(* IEC 61131-3 sources: STAR-PLC-Agent/results/raw/four_group_20261114/star_terra/PUB012/generation/sim_00, 1 file *)

(* ---- test_program.st ---- *)
PROGRAM PLC_PRG
VAR
 BenchStep : UDINT := 0;
 BenchCalls : UDINT := 0;
 BenchDone : BOOL := FALSE;
 BenchLastTime : TIME := T#0ms;
 BenchClockReady : BOOL := FALSE;
 BenchCurrentTime : TIME := T#0ms;
 TraceDt : ARRAY[0..15] OF UDINT;
 BenchUut0 : FB_Task;
 BenchUut1 : FB_Task;
 TraceIn_THICKNESS_FAULT : ARRAY[0..15] OF BOOL;
 TraceIn_THICKNESS_SIGNAL_VALID : ARRAY[0..15] OF BOOL;
 TraceIn_CUTTING_RUN : ARRAY[0..15] OF BOOL;
 TraceIn_FaultTimestamp : ARRAY[0..15] OF DINT;
 TraceIn_CycleTime : ARRAY[0..15] OF TIME;
 TraceOut_THICKNESS_ALARM : ARRAY[0..15] OF BOOL;
 TraceOut_Slab_Fault_Counter : ARRAY[0..15] OF UINT;
 TraceOut_Slab_Runtime_Accumulator : ARRAY[0..15] OF LTIME;
 TraceOut_Slab_Fault_History_0 : ARRAY[0..15] OF DINT;
 TraceOut_Slab_Fault_History_1 : ARRAY[0..15] OF DINT;
 TraceOut_Slab_Fault_History_2 : ARRAY[0..15] OF DINT;
 TraceOut_Slab_Fault_History_3 : ARRAY[0..15] OF DINT;
 TraceOut_Slab_Fault_History_4 : ARRAY[0..15] OF DINT;
END_VAR

IF NOT BenchDone THEN
 BenchCurrentTime := TIME();
 IF NOT BenchClockReady THEN
  BenchLastTime := BenchCurrentTime;
  BenchClockReady := TRUE;
 ELSE
 CASE BenchStep OF
 0:
  IF BenchCurrentTime - BenchLastTime >= UDINT_TO_TIME(10) THEN
   TraceDt[0] := TIME_TO_UDINT(BenchCurrentTime - BenchLastTime);
   BenchLastTime := BenchCurrentTime;
   BenchUut0.THICKNESS_FAULT := FALSE;
   BenchUut0.THICKNESS_SIGNAL_VALID := FALSE;
   BenchUut0.CUTTING_RUN := TRUE;
   BenchUut0.FaultTimestamp := DINT#0;
   BenchUut0.CycleTime := TIME#10ms;
   TraceIn_THICKNESS_FAULT[0] := BenchUut0.THICKNESS_FAULT;
   TraceIn_THICKNESS_SIGNAL_VALID[0] := BenchUut0.THICKNESS_SIGNAL_VALID;
   TraceIn_CUTTING_RUN[0] := BenchUut0.CUTTING_RUN;
   TraceIn_FaultTimestamp[0] := BenchUut0.FaultTimestamp;
   TraceIn_CycleTime[0] := BenchUut0.CycleTime;
   BenchUut0();
   TraceOut_THICKNESS_ALARM[0] := BenchUut0.THICKNESS_ALARM;
   TraceOut_Slab_Fault_Counter[0] := BenchUut0.Slab_Fault_Counter;
   TraceOut_Slab_Runtime_Accumulator[0] := BenchUut0.Slab_Runtime_Accumulator;
   TraceOut_Slab_Fault_History_0[0] := BenchUut0.Slab_Fault_History[0];
   TraceOut_Slab_Fault_History_1[0] := BenchUut0.Slab_Fault_History[1];
   TraceOut_Slab_Fault_History_2[0] := BenchUut0.Slab_Fault_History[2];
   TraceOut_Slab_Fault_History_3[0] := BenchUut0.Slab_Fault_History[3];
   TraceOut_Slab_Fault_History_4[0] := BenchUut0.Slab_Fault_History[4];
   BenchCalls := BenchCalls + 1;
   BenchStep := BenchStep + 1;
  END_IF;
 1:
  IF BenchCurrentTime - BenchLastTime >= UDINT_TO_TIME(100) THEN
   TraceDt[1] := TIME_TO_UDINT(BenchCurrentTime - BenchLastTime);
   BenchLastTime := BenchCurrentTime;
   BenchUut0.THICKNESS_FAULT := FALSE;
   BenchUut0.THICKNESS_SIGNAL_VALID := TRUE;
   BenchUut0.CUTTING_RUN := TRUE;
   BenchUut0.FaultTimestamp := DINT#0;
   BenchUut0.CycleTime := TIME#100ms;
   TraceIn_THICKNESS_FAULT[1] := BenchUut0.THICKNESS_FAULT;
   TraceIn_THICKNESS_SIGNAL_VALID[1] := BenchUut0.THICKNESS_SIGNAL_VALID;
   TraceIn_CUTTING_RUN[1] := BenchUut0.CUTTING_RUN;
   TraceIn_FaultTimestamp[1] := BenchUut0.FaultTimestamp;
   TraceIn_CycleTime[1] := BenchUut0.CycleTime;
   BenchUut0();
   TraceOut_THICKNESS_ALARM[1] := BenchUut0.THICKNESS_ALARM;
   TraceOut_Slab_Fault_Counter[1] := BenchUut0.Slab_Fault_Counter;
   TraceOut_Slab_Runtime_Accumulator[1] := BenchUut0.Slab_Runtime_Accumulator;
   TraceOut_Slab_Fault_History_0[1] := BenchUut0.Slab_Fault_History[0];
   TraceOut_Slab_Fault_History_1[1] := BenchUut0.Slab_Fault_History[1];
   TraceOut_Slab_Fault_History_2[1] := BenchUut0.Slab_Fault_History[2];
   TraceOut_Slab_Fault_History_3[1] := BenchUut0.Slab_Fault_History[3];
   TraceOut_Slab_Fault_History_4[1] := BenchUut0.Slab_Fault_History[4];
   BenchCalls := BenchCalls + 1;
   BenchStep := BenchStep + 1;
  END_IF;
 2:
  IF BenchCurrentTime - BenchLastTime >= UDINT_TO_TIME(20) THEN
   TraceDt[2] := TIME_TO_UDINT(BenchCurrentTime - BenchLastTime);
   BenchLastTime := BenchCurrentTime;
   BenchUut0.THICKNESS_FAULT := TRUE;
   BenchUut0.THICKNESS_SIGNAL_VALID := TRUE;
   BenchUut0.CUTTING_RUN := TRUE;
   BenchUut0.FaultTimestamp := DINT#101;
   BenchUut0.CycleTime := TIME#20ms;
   TraceIn_THICKNESS_FAULT[2] := BenchUut0.THICKNESS_FAULT;
   TraceIn_THICKNESS_SIGNAL_VALID[2] := BenchUut0.THICKNESS_SIGNAL_VALID;
   TraceIn_CUTTING_RUN[2] := BenchUut0.CUTTING_RUN;
   TraceIn_FaultTimestamp[2] := BenchUut0.FaultTimestamp;
   TraceIn_CycleTime[2] := BenchUut0.CycleTime;
   BenchUut0();
   TraceOut_THICKNESS_ALARM[2] := BenchUut0.THICKNESS_ALARM;
   TraceOut_Slab_Fault_Counter[2] := BenchUut0.Slab_Fault_Counter;
   TraceOut_Slab_Runtime_Accumulator[2] := BenchUut0.Slab_Runtime_Accumulator;
   TraceOut_Slab_Fault_History_0[2] := BenchUut0.Slab_Fault_History[0];
   TraceOut_Slab_Fault_History_1[2] := BenchUut0.Slab_Fault_History[1];
   TraceOut_Slab_Fault_History_2[2] := BenchUut0.Slab_Fault_History[2];
   TraceOut_Slab_Fault_History_3[2] := BenchUut0.Slab_Fault_History[3];
   TraceOut_Slab_Fault_History_4[2] := BenchUut0.Slab_Fault_History[4];
   BenchCalls := BenchCalls + 1;
   BenchStep := BenchStep + 1;
  END_IF;
 3:
  IF BenchCurrentTime - BenchLastTime >= UDINT_TO_TIME(600) THEN
   TraceDt[3] := TIME_TO_UDINT(BenchCurrentTime - BenchLastTime);
   BenchLastTime := BenchCurrentTime;
   BenchUut0.THICKNESS_FAULT := TRUE;
   BenchUut0.THICKNESS_SIGNAL_VALID := TRUE;
   BenchUut0.CUTTING_RUN := TRUE;
   BenchUut0.FaultTimestamp := DINT#999;
   BenchUut0.CycleTime := TIME#600ms;
   TraceIn_THICKNESS_FAULT[3] := BenchUut0.THICKNESS_FAULT;
   TraceIn_THICKNESS_SIGNAL_VALID[3] := BenchUut0.THICKNESS_SIGNAL_VALID;
   TraceIn_CUTTING_RUN[3] := BenchUut0.CUTTING_RUN;
   TraceIn_FaultTimestamp[3] := BenchUut0.FaultTimestamp;
   TraceIn_CycleTime[3] := BenchUut0.CycleTime;
   BenchUut0();
   TraceOut_THICKNESS_ALARM[3] := BenchUut0.THICKNESS_ALARM;
   TraceOut_Slab_Fault_Counter[3] := BenchUut0.Slab_Fault_Counter;
   TraceOut_Slab_Runtime_Accumulator[3] := BenchUut0.Slab_Runtime_Accumulator;
   TraceOut_Slab_Fault_History_0[3] := BenchUut0.Slab_Fault_History[0];
   TraceOut_Slab_Fault_History_1[3] := BenchUut0.Slab_Fault_History[1];
   TraceOut_Slab_Fault_History_2[3] := BenchUut0.Slab_Fault_History[2];
   TraceOut_Slab_Fault_History_3[3] := BenchUut0.Slab_Fault_History[3];
   TraceOut_Slab_Fault_History_4[3] := BenchUut0.Slab_Fault_History[4];
   BenchCalls := BenchCalls + 1;
   BenchStep := BenchStep + 1;
  END_IF;
 4:
  IF BenchCurrentTime - BenchLastTime >= UDINT_TO_TIME(1) THEN
   TraceDt[4] := TIME_TO_UDINT(BenchCurrentTime - BenchLastTime);
   BenchLastTime := BenchCurrentTime;
   BenchUut0.THICKNESS_FAULT := FALSE;
   BenchUut0.THICKNESS_SIGNAL_VALID := TRUE;
   BenchUut0.CUTTING_RUN := FALSE;
   BenchUut0.FaultTimestamp := DINT#999;
   BenchUut0.CycleTime := TIME#1ms;
   TraceIn_THICKNESS_FAULT[4] := BenchUut0.THICKNESS_FAULT;
   TraceIn_THICKNESS_SIGNAL_VALID[4] := BenchUut0.THICKNESS_SIGNAL_VALID;
   TraceIn_CUTTING_RUN[4] := BenchUut0.CUTTING_RUN;
   TraceIn_FaultTimestamp[4] := BenchUut0.FaultTimestamp;
   TraceIn_CycleTime[4] := BenchUut0.CycleTime;
   BenchUut0();
   TraceOut_THICKNESS_ALARM[4] := BenchUut0.THICKNESS_ALARM;
   TraceOut_Slab_Fault_Counter[4] := BenchUut0.Slab_Fault_Counter;
   TraceOut_Slab_Runtime_Accumulator[4] := BenchUut0.Slab_Runtime_Accumulator;
   TraceOut_Slab_Fault_History_0[4] := BenchUut0.Slab_Fault_History[0];
   TraceOut_Slab_Fault_History_1[4] := BenchUut0.Slab_Fault_History[1];
   TraceOut_Slab_Fault_History_2[4] := BenchUut0.Slab_Fault_History[2];
   TraceOut_Slab_Fault_History_3[4] := BenchUut0.Slab_Fault_History[3];
   TraceOut_Slab_Fault_History_4[4] := BenchUut0.Slab_Fault_History[4];
   BenchCalls := BenchCalls + 1;
   BenchStep := BenchStep + 1;
  END_IF;
 5:
  IF BenchCurrentTime - BenchLastTime >= UDINT_TO_TIME(20) THEN
   TraceDt[5] := TIME_TO_UDINT(BenchCurrentTime - BenchLastTime);
   BenchLastTime := BenchCurrentTime;
   BenchUut0.THICKNESS_FAULT := TRUE;
   BenchUut0.THICKNESS_SIGNAL_VALID := TRUE;
   BenchUut0.CUTTING_RUN := TRUE;
   BenchUut0.FaultTimestamp := DINT#202;
   BenchUut0.CycleTime := TIME#20ms;
   TraceIn_THICKNESS_FAULT[5] := BenchUut0.THICKNESS_FAULT;
   TraceIn_THICKNESS_SIGNAL_VALID[5] := BenchUut0.THICKNESS_SIGNAL_VALID;
   TraceIn_CUTTING_RUN[5] := BenchUut0.CUTTING_RUN;
   TraceIn_FaultTimestamp[5] := BenchUut0.FaultTimestamp;
   TraceIn_CycleTime[5] := BenchUut0.CycleTime;
   BenchUut0();
   TraceOut_THICKNESS_ALARM[5] := BenchUut0.THICKNESS_ALARM;
   TraceOut_Slab_Fault_Counter[5] := BenchUut0.Slab_Fault_Counter;
   TraceOut_Slab_Runtime_Accumulator[5] := BenchUut0.Slab_Runtime_Accumulator;
   TraceOut_Slab_Fault_History_0[5] := BenchUut0.Slab_Fault_History[0];
   TraceOut_Slab_Fault_History_1[5] := BenchUut0.Slab_Fault_History[1];
   TraceOut_Slab_Fault_History_2[5] := BenchUut0.Slab_Fault_History[2];
   TraceOut_Slab_Fault_History_3[5] := BenchUut0.Slab_Fault_History[3];
   TraceOut_Slab_Fault_History_4[5] := BenchUut0.Slab_Fault_History[4];
   BenchCalls := BenchCalls + 1;
   BenchStep := BenchStep + 1;
  END_IF;
 6:
  IF BenchCurrentTime - BenchLastTime >= UDINT_TO_TIME(10) THEN
   TraceDt[6] := TIME_TO_UDINT(BenchCurrentTime - BenchLastTime);
   BenchLastTime := BenchCurrentTime;
   BenchUut0.THICKNESS_FAULT := TRUE;
   BenchUut0.THICKNESS_SIGNAL_VALID := FALSE;
   BenchUut0.CUTTING_RUN := TRUE;
   BenchUut0.FaultTimestamp := DINT#250;
   BenchUut0.CycleTime := TIME#10ms;
   TraceIn_THICKNESS_FAULT[6] := BenchUut0.THICKNESS_FAULT;
   TraceIn_THICKNESS_SIGNAL_VALID[6] := BenchUut0.THICKNESS_SIGNAL_VALID;
   TraceIn_CUTTING_RUN[6] := BenchUut0.CUTTING_RUN;
   TraceIn_FaultTimestamp[6] := BenchUut0.FaultTimestamp;
   TraceIn_CycleTime[6] := BenchUut0.CycleTime;
   BenchUut0();
   TraceOut_THICKNESS_ALARM[6] := BenchUut0.THICKNESS_ALARM;
   TraceOut_Slab_Fault_Counter[6] := BenchUut0.Slab_Fault_Counter;
   TraceOut_Slab_Runtime_Accumulator[6] := BenchUut0.Slab_Runtime_Accumulator;
   TraceOut_Slab_Fault_History_0[6] := BenchUut0.Slab_Fault_History[0];
   TraceOut_Slab_Fault_History_1[6] := BenchUut0.Slab_Fault_History[1];
   TraceOut_Slab_Fault_History_2[6] := BenchUut0.Slab_Fault_History[2];
   TraceOut_Slab_Fault_History_3[6] := BenchUut0.Slab_Fault_History[3];
   TraceOut_Slab_Fault_History_4[6] := BenchUut0.Slab_Fault_History[4];
   BenchCalls := BenchCalls + 1;
   BenchStep := BenchStep + 1;
  END_IF;
 7:
  IF BenchCurrentTime - BenchLastTime >= UDINT_TO_TIME(10) THEN
   TraceDt[7] := TIME_TO_UDINT(BenchCurrentTime - BenchLastTime);
   BenchLastTime := BenchCurrentTime;
   BenchUut0.THICKNESS_FAULT := TRUE;
   BenchUut0.THICKNESS_SIGNAL_VALID := TRUE;
   BenchUut0.CUTTING_RUN := TRUE;
   BenchUut0.FaultTimestamp := DINT#303;
   BenchUut0.CycleTime := TIME#10ms;
   TraceIn_THICKNESS_FAULT[7] := BenchUut0.THICKNESS_FAULT;
   TraceIn_THICKNESS_SIGNAL_VALID[7] := BenchUut0.THICKNESS_SIGNAL_VALID;
   TraceIn_CUTTING_RUN[7] := BenchUut0.CUTTING_RUN;
   TraceIn_FaultTimestamp[7] := BenchUut0.FaultTimestamp;
   TraceIn_CycleTime[7] := BenchUut0.CycleTime;
   BenchUut0();
   TraceOut_THICKNESS_ALARM[7] := BenchUut0.THICKNESS_ALARM;
   TraceOut_Slab_Fault_Counter[7] := BenchUut0.Slab_Fault_Counter;
   TraceOut_Slab_Runtime_Accumulator[7] := BenchUut0.Slab_Runtime_Accumulator;
   TraceOut_Slab_Fault_History_0[7] := BenchUut0.Slab_Fault_History[0];
   TraceOut_Slab_Fault_History_1[7] := BenchUut0.Slab_Fault_History[1];
   TraceOut_Slab_Fault_History_2[7] := BenchUut0.Slab_Fault_History[2];
   TraceOut_Slab_Fault_History_3[7] := BenchUut0.Slab_Fault_History[3];
   TraceOut_Slab_Fault_History_4[7] := BenchUut0.Slab_Fault_History[4];
   BenchCalls := BenchCalls + 1;
   BenchStep := BenchStep + 1;
  END_IF;
 8:
  IF BenchCurrentTime - BenchLastTime >= UDINT_TO_TIME(1) THEN
   TraceDt[8] := TIME_TO_UDINT(BenchCurrentTime - BenchLastTime);
   BenchLastTime := BenchCurrentTime;
   BenchUut1.THICKNESS_FAULT := FALSE;
   BenchUut1.THICKNESS_SIGNAL_VALID := TRUE;
   BenchUut1.CUTTING_RUN := TRUE;
   BenchUut1.FaultTimestamp := DINT#0;
   BenchUut1.CycleTime := TIME#1ms;
   TraceIn_THICKNESS_FAULT[8] := BenchUut1.THICKNESS_FAULT;
   TraceIn_THICKNESS_SIGNAL_VALID[8] := BenchUut1.THICKNESS_SIGNAL_VALID;
   TraceIn_CUTTING_RUN[8] := BenchUut1.CUTTING_RUN;
   TraceIn_FaultTimestamp[8] := BenchUut1.FaultTimestamp;
   TraceIn_CycleTime[8] := BenchUut1.CycleTime;
   BenchUut1();
   TraceOut_THICKNESS_ALARM[8] := BenchUut1.THICKNESS_ALARM;
   TraceOut_Slab_Fault_Counter[8] := BenchUut1.Slab_Fault_Counter;
   TraceOut_Slab_Runtime_Accumulator[8] := BenchUut1.Slab_Runtime_Accumulator;
   TraceOut_Slab_Fault_History_0[8] := BenchUut1.Slab_Fault_History[0];
   TraceOut_Slab_Fault_History_1[8] := BenchUut1.Slab_Fault_History[1];
   TraceOut_Slab_Fault_History_2[8] := BenchUut1.Slab_Fault_History[2];
   TraceOut_Slab_Fault_History_3[8] := BenchUut1.Slab_Fault_History[3];
   TraceOut_Slab_Fault_History_4[8] := BenchUut1.Slab_Fault_History[4];
   BenchCalls := BenchCalls + 1;
   BenchStep := BenchStep + 1;
  END_IF;
 9:
  IF BenchCurrentTime - BenchLastTime >= UDINT_TO_TIME(1) THEN
   TraceDt[9] := TIME_TO_UDINT(BenchCurrentTime - BenchLastTime);
   BenchLastTime := BenchCurrentTime;
   BenchUut1.THICKNESS_FAULT := TRUE;
   BenchUut1.THICKNESS_SIGNAL_VALID := TRUE;
   BenchUut1.CUTTING_RUN := TRUE;
   BenchUut1.FaultTimestamp := DINT#-2147483648;
   BenchUut1.CycleTime := TIME#1ms;
   TraceIn_THICKNESS_FAULT[9] := BenchUut1.THICKNESS_FAULT;
   TraceIn_THICKNESS_SIGNAL_VALID[9] := BenchUut1.THICKNESS_SIGNAL_VALID;
   TraceIn_CUTTING_RUN[9] := BenchUut1.CUTTING_RUN;
   TraceIn_FaultTimestamp[9] := BenchUut1.FaultTimestamp;
   TraceIn_CycleTime[9] := BenchUut1.CycleTime;
   BenchUut1();
   TraceOut_THICKNESS_ALARM[9] := BenchUut1.THICKNESS_ALARM;
   TraceOut_Slab_Fault_Counter[9] := BenchUut1.Slab_Fault_Counter;
   TraceOut_Slab_Runtime_Accumulator[9] := BenchUut1.Slab_Runtime_Accumulator;
   TraceOut_Slab_Fault_History_0[9] := BenchUut1.Slab_Fault_History[0];
   TraceOut_Slab_Fault_History_1[9] := BenchUut1.Slab_Fault_History[1];
   TraceOut_Slab_Fault_History_2[9] := BenchUut1.Slab_Fault_History[2];
   TraceOut_Slab_Fault_History_3[9] := BenchUut1.Slab_Fault_History[3];
   TraceOut_Slab_Fault_History_4[9] := BenchUut1.Slab_Fault_History[4];
   BenchCalls := BenchCalls + 1;
   BenchStep := BenchStep + 1;
  END_IF;
 10:
  IF BenchCurrentTime - BenchLastTime >= UDINT_TO_TIME(499) THEN
   TraceDt[10] := TIME_TO_UDINT(BenchCurrentTime - BenchLastTime);
   BenchLastTime := BenchCurrentTime;
   BenchUut1.THICKNESS_FAULT := FALSE;
   BenchUut1.THICKNESS_SIGNAL_VALID := TRUE;
   BenchUut1.CUTTING_RUN := TRUE;
   BenchUut1.FaultTimestamp := DINT#0;
   BenchUut1.CycleTime := TIME#499ms;
   TraceIn_THICKNESS_FAULT[10] := BenchUut1.THICKNESS_FAULT;
   TraceIn_THICKNESS_SIGNAL_VALID[10] := BenchUut1.THICKNESS_SIGNAL_VALID;
   TraceIn_CUTTING_RUN[10] := BenchUut1.CUTTING_RUN;
   TraceIn_FaultTimestamp[10] := BenchUut1.FaultTimestamp;
   TraceIn_CycleTime[10] := BenchUut1.CycleTime;
   BenchUut1();
   TraceOut_THICKNESS_ALARM[10] := BenchUut1.THICKNESS_ALARM;
   TraceOut_Slab_Fault_Counter[10] := BenchUut1.Slab_Fault_Counter;
   TraceOut_Slab_Runtime_Accumulator[10] := BenchUut1.Slab_Runtime_Accumulator;
   TraceOut_Slab_Fault_History_0[10] := BenchUut1.Slab_Fault_History[0];
   TraceOut_Slab_Fault_History_1[10] := BenchUut1.Slab_Fault_History[1];
   TraceOut_Slab_Fault_History_2[10] := BenchUut1.Slab_Fault_History[2];
   TraceOut_Slab_Fault_History_3[10] := BenchUut1.Slab_Fault_History[3];
   TraceOut_Slab_Fault_History_4[10] := BenchUut1.Slab_Fault_History[4];
   BenchCalls := BenchCalls + 1;
   BenchStep := BenchStep + 1;
  END_IF;
 11:
  IF BenchCurrentTime - BenchLastTime >= UDINT_TO_TIME(1) THEN
   TraceDt[11] := TIME_TO_UDINT(BenchCurrentTime - BenchLastTime);
   BenchLastTime := BenchCurrentTime;
   BenchUut1.THICKNESS_FAULT := TRUE;
   BenchUut1.THICKNESS_SIGNAL_VALID := TRUE;
   BenchUut1.CUTTING_RUN := TRUE;
   BenchUut1.FaultTimestamp := DINT#2147483647;
   BenchUut1.CycleTime := TIME#1ms;
   TraceIn_THICKNESS_FAULT[11] := BenchUut1.THICKNESS_FAULT;
   TraceIn_THICKNESS_SIGNAL_VALID[11] := BenchUut1.THICKNESS_SIGNAL_VALID;
   TraceIn_CUTTING_RUN[11] := BenchUut1.CUTTING_RUN;
   TraceIn_FaultTimestamp[11] := BenchUut1.FaultTimestamp;
   TraceIn_CycleTime[11] := BenchUut1.CycleTime;
   BenchUut1();
   TraceOut_THICKNESS_ALARM[11] := BenchUut1.THICKNESS_ALARM;
   TraceOut_Slab_Fault_Counter[11] := BenchUut1.Slab_Fault_Counter;
   TraceOut_Slab_Runtime_Accumulator[11] := BenchUut1.Slab_Runtime_Accumulator;
   TraceOut_Slab_Fault_History_0[11] := BenchUut1.Slab_Fault_History[0];
   TraceOut_Slab_Fault_History_1[11] := BenchUut1.Slab_Fault_History[1];
   TraceOut_Slab_Fault_History_2[11] := BenchUut1.Slab_Fault_History[2];
   TraceOut_Slab_Fault_History_3[11] := BenchUut1.Slab_Fault_History[3];
   TraceOut_Slab_Fault_History_4[11] := BenchUut1.Slab_Fault_History[4];
   BenchCalls := BenchCalls + 1;
   BenchStep := BenchStep + 1;
  END_IF;
 12:
  IF BenchCurrentTime - BenchLastTime >= UDINT_TO_TIME(499) THEN
   TraceDt[12] := TIME_TO_UDINT(BenchCurrentTime - BenchLastTime);
   BenchLastTime := BenchCurrentTime;
   BenchUut1.THICKNESS_FAULT := FALSE;
   BenchUut1.THICKNESS_SIGNAL_VALID := TRUE;
   BenchUut1.CUTTING_RUN := TRUE;
   BenchUut1.FaultTimestamp := DINT#0;
   BenchUut1.CycleTime := TIME#499ms;
   TraceIn_THICKNESS_FAULT[12] := BenchUut1.THICKNESS_FAULT;
   TraceIn_THICKNESS_SIGNAL_VALID[12] := BenchUut1.THICKNESS_SIGNAL_VALID;
   TraceIn_CUTTING_RUN[12] := BenchUut1.CUTTING_RUN;
   TraceIn_FaultTimestamp[12] := BenchUut1.FaultTimestamp;
   TraceIn_CycleTime[12] := BenchUut1.CycleTime;
   BenchUut1();
   TraceOut_THICKNESS_ALARM[12] := BenchUut1.THICKNESS_ALARM;
   TraceOut_Slab_Fault_Counter[12] := BenchUut1.Slab_Fault_Counter;
   TraceOut_Slab_Runtime_Accumulator[12] := BenchUut1.Slab_Runtime_Accumulator;
   TraceOut_Slab_Fault_History_0[12] := BenchUut1.Slab_Fault_History[0];
   TraceOut_Slab_Fault_History_1[12] := BenchUut1.Slab_Fault_History[1];
   TraceOut_Slab_Fault_History_2[12] := BenchUut1.Slab_Fault_History[2];
   TraceOut_Slab_Fault_History_3[12] := BenchUut1.Slab_Fault_History[3];
   TraceOut_Slab_Fault_History_4[12] := BenchUut1.Slab_Fault_History[4];
   BenchCalls := BenchCalls + 1;
   BenchStep := BenchStep + 1;
  END_IF;
 13:
  IF BenchCurrentTime - BenchLastTime >= UDINT_TO_TIME(1) THEN
   TraceDt[13] := TIME_TO_UDINT(BenchCurrentTime - BenchLastTime);
   BenchLastTime := BenchCurrentTime;
   BenchUut1.THICKNESS_FAULT := FALSE;
   BenchUut1.THICKNESS_SIGNAL_VALID := TRUE;
   BenchUut1.CUTTING_RUN := TRUE;
   BenchUut1.FaultTimestamp := DINT#0;
   BenchUut1.CycleTime := TIME#1ms;
   TraceIn_THICKNESS_FAULT[13] := BenchUut1.THICKNESS_FAULT;
   TraceIn_THICKNESS_SIGNAL_VALID[13] := BenchUut1.THICKNESS_SIGNAL_VALID;
   TraceIn_CUTTING_RUN[13] := BenchUut1.CUTTING_RUN;
   TraceIn_FaultTimestamp[13] := BenchUut1.FaultTimestamp;
   TraceIn_CycleTime[13] := BenchUut1.CycleTime;
   BenchUut1();
   TraceOut_THICKNESS_ALARM[13] := BenchUut1.THICKNESS_ALARM;
   TraceOut_Slab_Fault_Counter[13] := BenchUut1.Slab_Fault_Counter;
   TraceOut_Slab_Runtime_Accumulator[13] := BenchUut1.Slab_Runtime_Accumulator;
   TraceOut_Slab_Fault_History_0[13] := BenchUut1.Slab_Fault_History[0];
   TraceOut_Slab_Fault_History_1[13] := BenchUut1.Slab_Fault_History[1];
   TraceOut_Slab_Fault_History_2[13] := BenchUut1.Slab_Fault_History[2];
   TraceOut_Slab_Fault_History_3[13] := BenchUut1.Slab_Fault_History[3];
   TraceOut_Slab_Fault_History_4[13] := BenchUut1.Slab_Fault_History[4];
   BenchCalls := BenchCalls + 1;
   BenchStep := BenchStep + 1;
  END_IF;
 14:
  IF BenchCurrentTime - BenchLastTime >= UDINT_TO_TIME(1) THEN
   TraceDt[14] := TIME_TO_UDINT(BenchCurrentTime - BenchLastTime);
   BenchLastTime := BenchCurrentTime;
   BenchUut1.THICKNESS_FAULT := TRUE;
   BenchUut1.THICKNESS_SIGNAL_VALID := TRUE;
   BenchUut1.CUTTING_RUN := TRUE;
   BenchUut1.FaultTimestamp := DINT#0;
   BenchUut1.CycleTime := TIME#1ms;
   TraceIn_THICKNESS_FAULT[14] := BenchUut1.THICKNESS_FAULT;
   TraceIn_THICKNESS_SIGNAL_VALID[14] := BenchUut1.THICKNESS_SIGNAL_VALID;
   TraceIn_CUTTING_RUN[14] := BenchUut1.CUTTING_RUN;
   TraceIn_FaultTimestamp[14] := BenchUut1.FaultTimestamp;
   TraceIn_CycleTime[14] := BenchUut1.CycleTime;
   BenchUut1();
   TraceOut_THICKNESS_ALARM[14] := BenchUut1.THICKNESS_ALARM;
   TraceOut_Slab_Fault_Counter[14] := BenchUut1.Slab_Fault_Counter;
   TraceOut_Slab_Runtime_Accumulator[14] := BenchUut1.Slab_Runtime_Accumulator;
   TraceOut_Slab_Fault_History_0[14] := BenchUut1.Slab_Fault_History[0];
   TraceOut_Slab_Fault_History_1[14] := BenchUut1.Slab_Fault_History[1];
   TraceOut_Slab_Fault_History_2[14] := BenchUut1.Slab_Fault_History[2];
   TraceOut_Slab_Fault_History_3[14] := BenchUut1.Slab_Fault_History[3];
   TraceOut_Slab_Fault_History_4[14] := BenchUut1.Slab_Fault_History[4];
   BenchCalls := BenchCalls + 1;
   BenchStep := BenchStep + 1;
  END_IF;
 15:
  IF BenchCurrentTime - BenchLastTime >= UDINT_TO_TIME(1) THEN
   TraceDt[15] := TIME_TO_UDINT(BenchCurrentTime - BenchLastTime);
   BenchLastTime := BenchCurrentTime;
   BenchUut1.THICKNESS_FAULT := FALSE;
   BenchUut1.THICKNESS_SIGNAL_VALID := TRUE;
   BenchUut1.CUTTING_RUN := FALSE;
   BenchUut1.FaultTimestamp := DINT#1;
   BenchUut1.CycleTime := TIME#1ms;
   TraceIn_THICKNESS_FAULT[15] := BenchUut1.THICKNESS_FAULT;
   TraceIn_THICKNESS_SIGNAL_VALID[15] := BenchUut1.THICKNESS_SIGNAL_VALID;
   TraceIn_CUTTING_RUN[15] := BenchUut1.CUTTING_RUN;
   TraceIn_FaultTimestamp[15] := BenchUut1.FaultTimestamp;
   TraceIn_CycleTime[15] := BenchUut1.CycleTime;
   BenchUut1();
   TraceOut_THICKNESS_ALARM[15] := BenchUut1.THICKNESS_ALARM;
   TraceOut_Slab_Fault_Counter[15] := BenchUut1.Slab_Fault_Counter;
   TraceOut_Slab_Runtime_Accumulator[15] := BenchUut1.Slab_Runtime_Accumulator;
   TraceOut_Slab_Fault_History_0[15] := BenchUut1.Slab_Fault_History[0];
   TraceOut_Slab_Fault_History_1[15] := BenchUut1.Slab_Fault_History[1];
   TraceOut_Slab_Fault_History_2[15] := BenchUut1.Slab_Fault_History[2];
   TraceOut_Slab_Fault_History_3[15] := BenchUut1.Slab_Fault_History[3];
   TraceOut_Slab_Fault_History_4[15] := BenchUut1.Slab_Fault_History[4];
   BenchCalls := BenchCalls + 1;
   BenchStep := BenchStep + 1;
  END_IF;
 END_CASE;
 END_IF;
 IF BenchStep >= 16 THEN BenchDone := TRUE; END_IF;
END_IF;
END_PROGRAM
